TYPE "ST_DeclarationCellHal"
VERSION : 0.1
   STRUCT
      "Clamp" {ExternalAccessible := 'False'; ExternalVisible := 'False'; ExternalWritable := 'False'} : "ST_DeclarationLeafHal";
      "Gate" {ExternalAccessible := 'False'; ExternalVisible := 'False'; ExternalWritable := 'False'} : "ST_DeclarationLeafHal";
   END_STRUCT;
END_TYPE
